(* IEC 61131-3 sources: 2026_Projet_YGO_ExcavatriceDragage/CODE_BACKUP/CODE_20260904_AvantWeekendBackup_v0.6.34/J_SUPERVISION/_TYPES/5_ASSISTANCE_DRAGAGE, 14 files *)

(* ---- ST_ChainDredgingAssist.st ---- *)
TYPE ST_ChainDredgingAssist :
STRUCT
    Idx101_EnableDiveSearch          : BOOL; // 1 = Assistance Plongée Armée (IHM) | 0 = Désarmée
    Idx102_EnableExtractionSequence  : BOOL; // 1 = Assistance Extraction Armée (IHM) | 0 = Désarmée
    Idx103_EnableDumpAtTremie        : BOOL; // 1 = Mode Vidage Trémie Armé (IHM) | 0 = Désarmé

    Idx201_DiveReady                 : BOOL; // 1 = Assistance Plongée Prête | 0 = Non Prête
    Idx202_DiveBusy                  : BOOL; // 1 = Séquence Plongée En Cours | 0 = Repos
    Idx203_DiveDone                  : BOOL; // 1 = Fond Confirmé | 0 = En Cours
    Idx204_DiveState                 : E_DiveSearchState; // État interne séquenceur plongée
    Idx205_DiveError                 : BOOL; // 0 = Sain | 1 = Défaut Plongée
    Idx206_DiveErrorId                : WORD; // bit0: préconditions, bit1: séquence Kobold, bit2: config seuils
    Idx207_BottomTouchConfirmed      : BOOL; // 1 = Contact Fond Confirmé (Kobold ou manuel) | 0 = Non Confirmé
    Idx208_DiveStepAtFault           : E_DiveSearchState; // Étape figée à l'apparition du défaut plongée (ERROR_HOLD masque l'état vivant)

    Idx301_ExtractionReady           : BOOL; // 1 = Assistance Extraction Prête | 0 = Non Prête
    Idx302_ExtractionBusy            : BOOL; // 1 = Séquence Extraction En Cours | 0 = Repos
    Idx303_ExtractionDone            : BOOL; // 1 = Extraction Terminée | 0 = En Cours
    Idx304_ExtractionState           : E_ExtractionAssistState; // État interne séquenceur extraction
    Idx305_ExtractionError           : BOOL; // 0 = Sain | 1 = Défaut Extraction
    Idx306_ExtractionErrorId          : WORD; // bit0: fond absent, bit1: fermeture, bit2: contrôle remontée, bit3: config
    Idx307_ExtractionStepAtFault     : E_ExtractionAssistState; // Étape figée à l'apparition du défaut extraction (ERROR_HOLD masque l'état vivant)

    Idx401_OperatorActionId          : WORD;       // Identifiant consigne opérateur conduite (0 = aucune)
    Idx402_OperatorAction            : STRING(120); // Texte consigne opérateur (secours affichage)

    Idx501_DumpAtTremieArmed         : BOOL; // 1 = Bit IHM TglEnableDumpAtTremie actif | 0 = Désarmé
    Idx502_DumpAtTremieAssistActive  : BOOL; // 1 = Mode réellement actif (armé ET Mode MAINT_N1/N2) | 0 = Inactif
    Idx503_DumpAtTremieAtTremie      : BOOL; // 1 = M3 à la position Trémie | 0 = Ailleurs
    Idx504_DumpAtTremieBucketOpenArmed : BOOL; // 1 = Ouverture benne armée par ce mode | 0 = Non armée
    Idx505_DumpAtTremieDescentLocked : BOOL; // 1 = Descending M1/M2 verrouillée (M3 hors P1/Maintenance) | 0 = Libre

    Idx601_BypassDiveActive          : BOOL; // 1 = Bypass séquence DiveSearch armé (IHM)
    Idx602_BypassKoboldBottomTouched : BOOL; // 1 = Fond confirmé par le bypass (front montant Kobold en descente)
END_STRUCT
END_TYPE

(* ---- ST_CycleAssistToggles.st ---- *)
(* ═══════════════════════════════════════════════════════════════
   🎛️ ST_CycleAssistToggles — Toggles assistance mémorisés au boot
   📄 Doc : DOC/AF/AF_Partie-04_Mode_SemiAuto_Sequenceur_v2.3.md §3ter
   ═══════════════════════════════════════════════════════════════ *)
TYPE ST_CycleAssistToggles :
STRUCT
    TglEnableDiveSearch         : BOOL := FALSE; (* Mode assistance plongée mémorisé *)
    TglEnableExtractionSequence : BOOL := FALSE; (* Mode assistance extraction mémorisé *)
    TglEnableDumpAtTremie       : BOOL := FALSE; (* Mode assistance vidage trémie mémorisé *)
    Initialized                 : BOOL := FALSE; (* 🚦 flag restauration boot *)
END_STRUCT
END_TYPE

(* ---- ST_CycleDiveSearchCfg.st ---- *)
(* ═══════════════════════════════════════════════════════════════
   ⚙️ ST_CycleDiveSearchCfg — Réglages persistants cycle plongée (DiveSearch)
   📄 Doc : DOC/AF/AF_Partie-04_Mode_SemiAuto_Sequenceur_v2.3.md §3ter
   ═══════════════════════════════════════════════════════════════ *)
TYPE ST_CycleDiveSearchCfg :
STRUCT
    DiveStartMin_M   : REAL := 1.0;  (* Position mini M1/M2 avant plongée *)
    ImmersionUpper_M : REAL := 0.5;  (* Borne haute fenêtre front immersion *)
    ImmersionLower_M : REAL := -0.5; (* Borne basse fenêtre front immersion *)
    Initialized      : BOOL := FALSE; (* 🚦 flag restauration boot *)
END_STRUCT
END_TYPE

(* ---- ST_CycleDiveSearchCmd.st ---- *)
(* ═══════════════════════════════════════════════════════════════
   🎮 ST_CycleDiveSearchCmd — Sélections IHM cycle plongée (DiveSearch)
   ═══════════════════════════════════════════════════════════════ *)
TYPE ST_CycleDiveSearchCmd :
STRUCT
    TglEnableDiveSearch         : BOOL := FALSE; (* Assistance plongée active *)
    TglBypassDiveSearchSequence : BOOL := FALSE; (* Bypass séquence DiveSearch *)
    TglBucketAtBottomConfirmed  : BOOL := FALSE; (* Attestation manuelle fond *)
END_STRUCT
END_TYPE

(* ---- ST_CycleDiveSearchHMI.st ---- *)
(* ═══════════════════════════════════════════════════════════════
   🪨 ST_CycleDiveSearchHMI — Échange IHM cycle plongée (DiveSearch)
   ═══════════════════════════════════════════════════════════════ *)
TYPE ST_CycleDiveSearchHMI :
STRUCT
    Cmd   : ST_CycleDiveSearchCmd;
    State : ST_CycleDiveSearchState;
    Cfg   : ST_CycleDiveSearchCfg;
END_STRUCT
END_TYPE

(* ---- ST_CycleDiveSearchState.st ---- *)
(* ═══════════════════════════════════════════════════════════════
   🚦 ST_CycleDiveSearchState — États publics cycle plongée (DiveSearch)
   ═══════════════════════════════════════════════════════════════ *)
TYPE ST_CycleDiveSearchState :
STRUCT
    DiveReady             : BOOL;
    DiveBusy              : BOOL;
    DiveDone              : BOOL;
    DiveError             : BOOL;
    DiveErrorId           : WORD;
    DiveState             : E_DiveSearchState;
    DiveStepAtFault       : E_DiveSearchState;
    BottomTouchConfirmed  : BOOL;
    BypassDiveActive      : BOOL; (* TglBypassDiveSearchSequence armé (descente couplée en cours) *)
    BypassKoboldBottomTouched : BOOL; (* Fond confirmé par le bypass (front montant Kobold en descente) *)
    OperatorActionId         : WORD;       (* Une seule consigne conduite, arbitré en PRG_03 *)
    OperatorAction           : STRING(120); (* Texte de secours ; IHM peut mapper l'identifiant *)
END_STRUCT
END_TYPE

(* ---- ST_CycleDumpAtTremieCfg.st ---- *)
(* ═══════════════════════════════════════════════════════════════
   ⚙️ ST_CycleDumpAtTremieCfg — Réglages persistants cycle vidage trémie (legacy)
   ═══════════════════════════════════════════════════════════════ *)
TYPE ST_CycleDumpAtTremieCfg :
STRUCT
    Initialized : BOOL := FALSE; (* 🚦 flag restauration boot *)
END_STRUCT
END_TYPE

(* ---- ST_CycleDumpAtTremieCmd.st ---- *)
(* ═══════════════════════════════════════════════════════════════
   🎮 ST_CycleDumpAtTremieCmd — Sélections IHM cycle vidage trémie (legacy)
   ═══════════════════════════════════════════════════════════════ *)
TYPE ST_CycleDumpAtTremieCmd :
STRUCT
    TglEnableDumpAtTremie : BOOL := FALSE; (* Mode vidage à la trémie — RESTREINT des mouvements dès le boot *)
END_STRUCT
END_TYPE

(* ---- ST_CycleDumpAtTremieHMI.st ---- *)
(* ═══════════════════════════════════════════════════════════════
   🪨 ST_CycleDumpAtTremieHMI — Échange IHM cycle vidage trémie (legacy)
   ═══════════════════════════════════════════════════════════════ *)
TYPE ST_CycleDumpAtTremieHMI :
STRUCT
    Cmd   : ST_CycleDumpAtTremieCmd;
    State : ST_CycleDumpAtTremieState;
    Cfg   : ST_CycleDumpAtTremieCfg;
END_STRUCT
END_TYPE

(* ---- ST_CycleDumpAtTremieState.st ---- *)
(* ═══════════════════════════════════════════════════════════════
   🚦 ST_CycleDumpAtTremieState — États publics cycle vidage trémie (legacy)
   ═══════════════════════════════════════════════════════════════ *)
TYPE ST_CycleDumpAtTremieState :
STRUCT
    DumpAtTremieArmed           : BOOL; (* TglEnableDumpAtTremie (bit IHM brut) *)
    DumpAtTremieAssistActive    : BOOL; (* Armé ET Mode MAINT_N1/N2 (mode réellement actif) *)
    DumpAtTremieAtTremie        : BOOL; (* M3_AtTremieStable *)
    DumpAtTremieBucketOpenArmed : BOOL; (* CmdOpen_IHM déclenché par ce mode *)
    DumpAtTremieDescentLocked   : BOOL; (* DescendPermit M1/M2 forcé par ce mode (hors P1/Maintenance) *)
END_STRUCT
END_TYPE

(* ---- ST_CycleExtractionCfg.st ---- *)
(* ═══════════════════════════════════════════════════════════════
   ⚙️ ST_CycleExtractionCfg — Réglages persistants cycle extraction
   📄 Doc : DOC/AF/AF_Partie-04_Mode_SemiAuto_Sequenceur_v2.3.md §3ter
   ═══════════════════════════════════════════════════════════════ *)
TYPE ST_CycleExtractionCfg :
STRUCT
    ExtractionControlDistance_M : REAL := 2.0; (* Remontée palier 1 avant accélération *)
    Initialized                 : BOOL := FALSE; (* 🚦 flag restauration boot *)
END_STRUCT
END_TYPE

(* ---- ST_CycleExtractionCmd.st ---- *)
(* ═══════════════════════════════════════════════════════════════
   🎮 ST_CycleExtractionCmd — Sélections IHM cycle extraction
   ═══════════════════════════════════════════════════════════════ *)
TYPE ST_CycleExtractionCmd :
STRUCT
    TglEnableExtractionSequence : BOOL := FALSE; (* Assistance extraction active *)
END_STRUCT
END_TYPE

(* ---- ST_CycleExtractionHMI.st ---- *)
(* ═══════════════════════════════════════════════════════════════
   🪨 ST_CycleExtractionHMI — Échange IHM cycle extraction
   ═══════════════════════════════════════════════════════════════ *)
TYPE ST_CycleExtractionHMI :
STRUCT
    Cmd   : ST_CycleExtractionCmd;
    State : ST_CycleExtractionState;
    Cfg   : ST_CycleExtractionCfg;
END_STRUCT
END_TYPE

(* ---- ST_CycleExtractionState.st ---- *)
(* ═══════════════════════════════════════════════════════════════
   🚦 ST_CycleExtractionState — États publics cycle extraction
   ═══════════════════════════════════════════════════════════════ *)
TYPE ST_CycleExtractionState :
STRUCT
    ExtractionReady       : BOOL;
    ExtractionBusy        : BOOL;
    ExtractionDone        : BOOL;
    ExtractionError       : BOOL;
    ExtractionErrorId     : WORD;
    ExtractionState       : E_ExtractionAssistState;
    ExtractionStepAtFault : E_ExtractionAssistState;
END_STRUCT
END_TYPE
